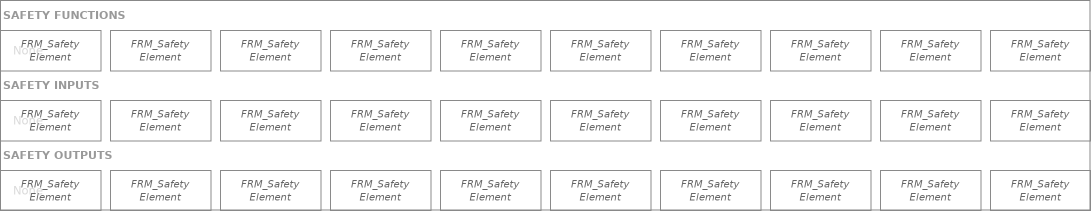
VISUALIZATION FRM_SafetyElementTable  // 1091x211
VAR_INPUT
    nFunctionCount: USINT;
    nInputCount: USINT; 
    nOutputCount: USINT;
END_VAR
    Label (10,30 91x41), "None"
    Label (10,100 91x41), "None"
    Label (10,170 91x41), "None"
    Frame (0,30 101x41), invisible if: nFunctionCount < 1
        shows FRM_SafetyElement(nIndex := 1, nOffset := 0)
    Frame (110,30 101x41), invisible if: nFunctionCount < 2
        shows FRM_SafetyElement(nIndex := 2, nOffset := 0)
    Label (0,0 161x31), "SAFETY FUNCTIONS"
    Label (0,70 161x31), "SAFETY INPUTS"
    Frame (0,100 101x41), invisible if: nInputCount < 1
        shows FRM_SafetyElement(nIndex := 1, nOffset := GVL_APP.nOFFSET_SAFE_INPUTS)
    Label (0,140 161x31)
    Frame (0,170 101x41), invisible if: nOutputCount < 1
        shows FRM_SafetyElement(nIndex := 1, nOffset := GVL_APP.nOFFSET_SAFE_OUTPUTS)
    Frame (110,170 101x41), invisible if: nOutputCount < 2
        shows FRM_SafetyElement(nIndex := 2, nOffset := GVL_APP.nOFFSET_SAFE_OUTPUTS)
    Frame (220,170 101x41), invisible if: nOutputCount < 3
        shows FRM_SafetyElement(nIndex := 3, nOffset := GVL_APP.nOFFSET_SAFE_OUTPUTS)
    Frame (110,100 101x41), invisible if: nInputCount < 2
        shows FRM_SafetyElement(nIndex := 2, nOffset := GVL_APP.nOFFSET_SAFE_INPUTS)
    Frame (220,30 101x41), invisible if: nFunctionCount < 3
        shows FRM_SafetyElement(nIndex := 3, nOffset := 0)
    Frame (330,30 101x41), invisible if: nFunctionCount < 4
        shows FRM_SafetyElement(nIndex := 4, nOffset := 0)
    Frame (440,30 101x41), invisible if: nFunctionCount < 5
        shows FRM_SafetyElement(nIndex := 5, nOffset := 0)
    Frame (550,30 101x41), invisible if: nFunctionCount < 6
        shows FRM_SafetyElement(nIndex := 6, nOffset := 0)
    Frame (660,30 101x41), invisible if: nFunctionCount < 7
        shows FRM_SafetyElement(nIndex := 7, nOffset := 0)
    Frame (770,30 101x41), invisible if: nFunctionCount < 8
        shows FRM_SafetyElement(nIndex := 8, nOffset := 0)
    Frame (880,30 101x41), invisible if: nFunctionCount < 9
        shows FRM_SafetyElement(nIndex := 9, nOffset := 0)
    Frame (220,100 101x41), invisible if: nInputCount < 3
        shows FRM_SafetyElement(nIndex := 3, nOffset := GVL_APP.nOFFSET_SAFE_INPUTS)
    Frame (330,100 101x41), invisible if: nInputCount < 4
        shows FRM_SafetyElement(nIndex := 4, nOffset := GVL_APP.nOFFSET_SAFE_INPUTS)
    Frame (440,100 101x41), invisible if: nInputCount < 5
        shows FRM_SafetyElement(nIndex := 5, nOffset := GVL_APP.nOFFSET_SAFE_INPUTS)
    Frame (550,100 101x41), invisible if: nInputCount < 6
        shows FRM_SafetyElement(nIndex := 6, nOffset := GVL_APP.nOFFSET_SAFE_INPUTS)
    Frame (660,100 101x41), invisible if: nInputCount < 7
        shows FRM_SafetyElement(nIndex := 7, nOffset := GVL_APP.nOFFSET_SAFE_INPUTS)
    Frame (770,100 101x41), invisible if: nInputCount < 8
        shows FRM_SafetyElement(nIndex := 8, nOffset := GVL_APP.nOFFSET_SAFE_INPUTS)
    Frame (880,100 101x41), invisible if: nInputCount < 9
        shows FRM_SafetyElement(nIndex := 9, nOffset := GVL_APP.nOFFSET_SAFE_INPUTS)
    Frame (990,100 101x41), invisible if: nInputCount < 10
        shows FRM_SafetyElement(nIndex := 10, nOffset := GVL_APP.nOFFSET_SAFE_INPUTS)
    Frame (330,170 101x41), invisible if: nOutputCount < 4
        shows FRM_SafetyElement(nIndex := 4, nOffset := GVL_APP.nOFFSET_SAFE_OUTPUTS)
    Frame (440,170 101x41), invisible if: nOutputCount < 5
        shows FRM_SafetyElement(nIndex := 5, nOffset := GVL_APP.nOFFSET_SAFE_OUTPUTS)
    Frame (550,170 101x41), invisible if: nOutputCount < 6
        shows FRM_SafetyElement(nIndex := 6, nOffset := GVL_APP.nOFFSET_SAFE_OUTPUTS)
    Frame (660,170 101x41), invisible if: nOutputCount < 7
        shows FRM_SafetyElement(nIndex := 7, nOffset := GVL_APP.nOFFSET_SAFE_OUTPUTS)
    Frame (770,170 101x41), invisible if: nOutputCount < 8
        shows FRM_SafetyElement(nIndex := 8, nOffset := GVL_APP.nOFFSET_SAFE_OUTPUTS)
    Frame (880,170 101x41), invisible if: nOutputCount < 9
        shows FRM_SafetyElement(nIndex := 9, nOffset := GVL_APP.nOFFSET_SAFE_OUTPUTS)
    Frame (990,170 101x41), invisible if: nOutputCount < 10
        shows FRM_SafetyElement(nIndex := 10, nOffset := GVL_APP.nOFFSET_SAFE_OUTPUTS)
    Frame (990,30 101x41), invisible if: nFunctionCount < 10
        shows FRM_SafetyElement(nIndex := 10, nOffset := 0)
    Label (0,140 161x31), "SAFETY OUTPUTS"
END_VISUALIZATION

(* stored: Version 1.1.0.1
   Visu FRM_SafetyElementTable: Id {2b1ae4e0-da87-0cb8-1607-3398f301c06a} *)
